// TIA Portal V21 export
// export: Created 2026-08-21T20:18:52.0075411Z, ExportSetting None, DisplayName Totally Integrated Automation Portal, DisplayVersion V21, DisplayName STEP 7 Professional, DisplayVersion V21, DisplayName STEP 7 Safety, DisplayVersion V21, DisplayName Tech WebApplication, DisplayVersion V21, DisplayName WinCC Basic/Comfort/Advanced, DisplayVersion V21, DisplayName WinCC Professional, DisplayVersion V21, DisplayName WinCC Unified, DisplayVersion V21
DATA_BLOCK "ReportValues_DB"   // DB35
AUTHOR : Siemens AG
FAMILY : ServiceControl
VERSION : 1.0
// stored: InstanceOfName ReportValues, InstanceOfType FB
"ReportValues"
   // VAR
   //    MTPAnalog { S7_SetPoint := 'True'} : Array[0..1] of "UDT_MTP_AnaReportValue";
   //    MTPDigital { S7_SetPoint := 'True'} : Array[0..0] of "UDT_MTP_DIntReportValue";
   //    MTPBinary { S7_SetPoint := 'True'} : Array[0..0] of "UDT_MTP_BinReportValue";
   //    MTPString { S7_SetPoint := 'True'} : Array[0..0] of "UDT_MTP_StringReportValue";
   // END_VAR
BEGIN
   MTPAnalog[0..1].V := 0.0;
   MTPAnalog[0..1].VSclMin := 0.0;
   MTPAnalog[0].VSclMax := 32.0;
   MTPAnalog[1].VSclMax := 100000.0;
   MTPAnalog[0].VUnit := 1351;
   MTPAnalog[1].VUnit := 1038;
END_DATA_BLOCK
